(* IEC 61131-3 sources: avi-aoi-management/scripts/ai-eval/ngau-nhien/kho/st-ud6-nhiet-on-off/mau/src, 2 files *)

(* ---- DieuKhienNhietLo.st ---- *)
FUNCTION_BLOCK DieuKhienNhietLo
VAR_INPUT
    BAT : BOOL;
    NHIET : REAL;
    SP : REAL;
    TRE : REAL;
    NGUONG_CAO : REAL;
    NGUONG_HH : REAL;
    RESET : BOOL;
END_VAR
VAR_OUTPUT
    SUOI : BOOL;
    CANH_BAO_CAO : BOOL;
    NGAT_HH : BOOL;
    LOI_CAM_BIEN : BOOL;
    TRANG_THAI : INT;  (* 0 TAT, 1 DIEU_KHIEN, 2 NGAT_HH, 3 LOI_CAM_BIEN *)
END_VAR
VAR
    boTre : TreHaiNguong;
END_VAR
    LOI_CAM_BIEN := NHIET < -50.0 OR NHIET > 500.0;
    boTre(X := NHIET, SP := SP, TRE := TRE);
    CANH_BAO_CAO := NOT LOI_CAM_BIEN AND NHIET >= NGUONG_CAO;
    IF NOT LOI_CAM_BIEN AND NHIET >= NGUONG_HH THEN
        NGAT_HH := TRUE;
    ELSIF RESET AND NOT LOI_CAM_BIEN AND NHIET < SP THEN
        NGAT_HH := FALSE;
    END_IF
    SUOI := BAT AND boTre.Q AND NOT NGAT_HH AND NOT LOI_CAM_BIEN;
    IF LOI_CAM_BIEN THEN
        TRANG_THAI := 3;
    ELSIF NGAT_HH THEN
        TRANG_THAI := 2;
    ELSIF NOT BAT THEN
        TRANG_THAI := 0;
    ELSE
        TRANG_THAI := 1;
    END_IF
END_FUNCTION_BLOCK

(* ---- TreHaiNguong.st ---- *)
FUNCTION_BLOCK TreHaiNguong
VAR_INPUT
    X : REAL;
    SP : REAL;
    TRE : REAL;
END_VAR
VAR_OUTPUT
    Q : BOOL;
END_VAR
    IF X <= SP - TRE THEN
        Q := TRUE;
    ELSIF X >= SP + TRE THEN
        Q := FALSE;
    END_IF
END_FUNCTION_BLOCK
